FUNCTION F_OPC_REMOTE (* OPC-UA-ID fuer einen Knoten auf einer anderen Station: opc_ua[ACTION;ENDPOINT#;NODE] *)
  (* Standard: 61499-1; Description: Copyright (c) 2026 Meisterschulen am Ostbahnhof This program and the accompanying materials are made available under the terms of the Eclipse Public License 2.0 which is available at https://www.eclipse.org/legal/epl-2.0/ SPDX-License-Identifier: EPL-2.0 *)
  (* Version 1.0, 2026-10-17, Franz Höpfinger, Meisterschulen am Ostbahnhof, initial implementation *)
  PACKAGE MyLib_OPC;
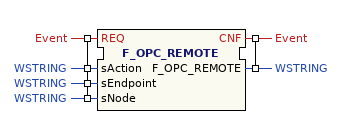
  EVENT_INPUT
    REQ WITH sAction, sEndpoint, sNode;
  END_EVENT
  EVENT_OUTPUT
    CNF WITH F_OPC_REMOTE;
  END_EVENT
  VAR_INPUT
    sAction : WSTRING; (* ACTION, z.B. WRITE oder CALL_METHOD *)
    sEndpoint : WSTRING; (* Endpunkt, z.B. opc.tcp://192.168.1.12:4840 *)
    sNode : WSTRING; (* Knoten, z.B. /Objects/X/Y,1:s=Y *)
  END_VAR
  VAR_OUTPUT
    F_OPC_REMOTE : WSTRING;
  END_VAR
  BODY IN ST:
PACKAGE MyLib_OPC;

(* OPC-UA-ID fuer einen Knoten auf einer anderen Station: opc_ua[ACTION;ENDPOINT#;NODE] *)
FUNCTION F_OPC_REMOTE : WSTRING

VAR_INPUT
	sAction : WSTRING; // ACTION, z.B. WRITE oder CALL_METHOD
	sEndpoint : WSTRING; // Endpunkt, z.B. opc.tcp://192.168.1.12:4840
	sNode : WSTRING; // Knoten, z.B. /Objects/X/Y,1:s=Y
END_VAR

F_OPC_REMOTE := CONCAT("opc_ua[", sAction, ";", sEndpoint, "#;", sNode, "]");

END_FUNCTION
  END_BODY
END_FUNCTION
